// TIA Portal V21 export
// export: Created 2026-11-07T17:04:58.1383967Z, ExportSetting WithDefaults, DisplayName Totally Integrated Automation Portal, DisplayVersion V21, DisplayName STEP 7 Professional, DisplayVersion V21, DisplayName STEP 7 Safety, DisplayVersion V21, DisplayName Tech WebApplication, DisplayVersion V21, DisplayName WinCC Basic/Comfort/Advanced, DisplayVersion V21, DisplayName WinCC Unified, DisplayVersion V21
TagTable "Default tag table"
  time : Real  (HMI_Connection_1, 1 s)
  P_SwOn : Bool  (HMI_Connection_1, 1 s)
